// TIA Portal V21 export
// export: Created 2026-11-18T10:00:00.0000000Z, ExportSetting None
ORGANIZATION_BLOCK "OB_Cyclic"   // OB30, LAD, CyclicInterrupt
{ S7_Optimized_Access := 'TRUE' }
// stored: CyclicTime 100000, PhaseOffset 0, SetENOAutomatically false
   VAR_INPUT
      Initial_Call : Bool;
      Event_Count : Int;
   END_VAR
   VAR_TEMP
      Tmp : Int;
   END_VAR
BEGIN

REGION Network 1: Cycle counter
   // counts by two unless held
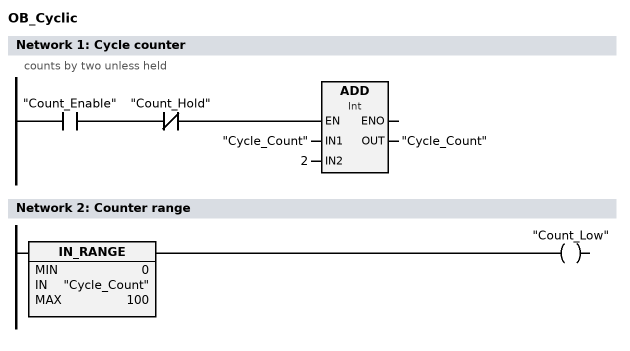
   RUNG wire#powerrail
      Contact( "Count_Enable" )
      I_Contact( "Count_Hold" )
      { S7_Templates := "SrcType := Int" } Add(in1 := "Cycle_Count", in2 := 2, out => "Cycle_Count")
   END_RUNG
   // the same network as SCL:
   IF "Count_Enable" AND NOT "Count_Hold" THEN "Cycle_Count" := "Cycle_Count" + 2; END_IF;
END_REGION

REGION Network 2: Counter range
   RUNG wire#powerrail
      { S7_Templates := "SrcType := Int" } InRange(min := 0, in := "Cycle_Count", max := 100)
      Coil( "Count_Low" )
   END_RUNG
   // the same network as SCL:
   "Count_Low" := (0 <= "Cycle_Count") AND ("Cycle_Count" <= 100);
END_REGION
END_ORGANIZATION_BLOCK
